{attribute 'Tc2GvlVarNames'}
VAR_GLOBAL
	(*fbCheckDivRealInfo: FB_CheckDivRealInfo;*)
END_VAR

(* stored: Version 1.1.0.1, ProductVersion 3.1.4024.15
   GVL GVL_FB_CheckDivRealInfo: Id {20bd6a95-3ab1-4313-bcde-363cfa647886} *)
